// TIA Portal V20 export
// export: Created 2026-10-12T05:42:31.3498917Z, ExportSetting WithDefaults, DisplayName Totally Integrated Automation Portal, DisplayVersion V20, DisplayName TIA Portal Openness, DisplayVersion V20, DisplayName TIA Portal Teamcenter Gateway, DisplayVersion V20, DisplayName TIA Portal Version Control Interface, DisplayVersion V20, DisplayName SINAMICS Startdrive Advanced, DisplayVersion V20 SP1 Update 2, DisplayName SINAMICS Startdrive G110M, G120, G120C, G120D, G120P, G115D, DisplayVersion V20 SP1 Update 2, DisplayName SINAMICS Startdrive G130, G150, S120, S150, SINAMICS MV, G220, S200, S210, DisplayVersion V20 SP1 Update 2, DisplayName STEP 7 Professional, DisplayVersion V20, DisplayName STEP 7 Safety, DisplayVersion V20, DisplayName WinCC Basic/Comfort/Advanced, DisplayVersion V20, DisplayName WinCC Professional, DisplayVersion V20, DisplayName WinCC Unified, DisplayVersion V20
FUNCTION "FRK_DecisionTake" : Int   // FC92, SCL
{ S7_Optimized_Access := 'TRUE' }
VERSION : 0.1
// stored: AutoNumber true, IsIECCheckEnabled false, SetENOAutomatically false, UDAEnableTagReadback false
   VAR_INPUT
      Owner : DInt;
   END_VAR
   VAR_IN_OUT
      AlarmLog : "FRK_AlarmLog";
   END_VAR
   VAR_TEMP
      Slot : Int;
   END_VAR
BEGIN

   #FRK_DecisionTake := 0;
   #Slot := "FRK_DecisionRoot"(Owner := #Owner, Create := FALSE);
   IF #Slot = 0 THEN
       RETURN;
   END_IF;
   IF "FRK_Decisions".Slots[#Slot].Owner <> #Owner THEN
       RETURN;
   END_IF;
   IF "FRK_Decisions".Slots[#Slot].Answer = 0 THEN
       RETURN;
   END_IF;
   #FRK_DecisionTake := "FRK_Decisions".Slots[#Slot].Answer;
   IF NOT "FRK_Decisions".Slots[#Slot].ResolutionLogged THEN
       "FRK_DecisionAudit"(AlarmLog := #AlarmLog,
                           Key := WSTRING#'std.audit.decisionOperatorResolved',
                           SourcePath := "FRK_Decisions".Slots[#Slot].Request.SourcePath,
                           Option := #FRK_DecisionTake);
   END_IF;
   "FRK_DecisionClear"(Slot := "FRK_Decisions".Slots[#Slot]);
END_FUNCTION
